// TIA Portal V21 export
// export: Created 2026-11-10T19:43:15.1099437Z, ExportSetting WithDefaults, DisplayName Totally Integrated Automation Portal, DisplayVersion V21 Update 3, DisplayName STEP 7 Professional, DisplayVersion V21 Update 3, DisplayName STEP 7 Safety, DisplayVersion V21, DisplayName Tech WebApplication, DisplayVersion V21, DisplayName WinCC Basic/Comfort/Advanced, DisplayVersion V21 Update 3, DisplayName WinCC Unified, DisplayVersion V21 Update 3
FUNCTION_BLOCK "FB_LadStruct"   // FB116, LAD
{ S7_Optimized_Access := 'TRUE' }
VERSION : 0.1
// stored: AutoNumber true, IsIECCheckEnabled false, IsRetainMemResEnabled false, MemoryReserve 100, SetENOAutomatically false, UDAEnableTagReadback false
   VAR_INPUT
      "a" : Bool;
      "b" : Bool;
      c : Bool;
      ia : Int;
   END_VAR
   VAR_OUTPUT
      q : Bool;
      q2 : Bool;
      io : Int;
      io2 : Int;
   END_VAR
   VAR
      ifc1 { S7_SetPoint := 'True'} : "FB_Iface";
      ton1 { S7_SetPoint := 'True'} : TON_TIME;
   END_VAR
BEGIN

REGION Network 1: Parallel branch
   // Branch with a second contact
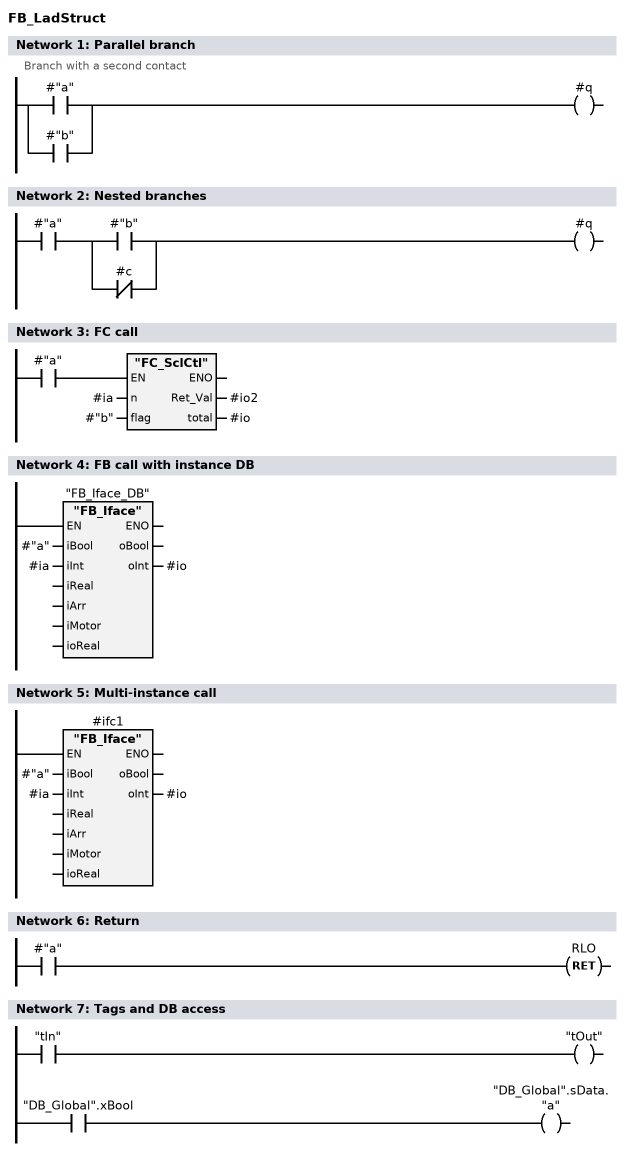
   RUNG wire#powerrail
      Contact( #"a" )
      wire#w1
      Coil( #q )
   END_RUNG
   RUNG wire#powerrail
      Contact( #"b" )
   END_RUNG wire#w1
   // the same network as SCL:
   #q := #"a" OR #"b";
END_REGION

REGION Network 2: Nested branches
   RUNG wire#powerrail
      Contact( #"a" )
      wire#w1
      Contact( #"b" )
      wire#w2
      Coil( #q )
   END_RUNG
   RUNG wire#w1
      I_Contact( #c )
   END_RUNG wire#w2
   // the same network as SCL:
   #q := #"a" AND (#"b" OR NOT #c);
END_REGION

REGION Network 3: FC call
   RUNG wire#powerrail
      Contact( #"a" )
      "FC_SclCtl"(n := #ia, flag := #"b", total => #io, Ret_Val => #io2)
   END_RUNG
   // the same network as SCL:
   IF #"a" THEN #io2 := "FC_SclCtl"(n := #ia, flag := #"b", total => #io); END_IF;
END_REGION

REGION Network 4: FB call with instance DB
   RUNG wire#powerrail
      "FB_Iface_DB"(iBool := #"a", iInt := #ia, oInt => #io, iReal :=, iArr :=, iMotor :=, oBool =>, ioReal :=)
   END_RUNG
   // the same network as SCL:
   "FB_Iface_DB"(iBool := #"a", iInt := #ia, oInt => #io);   // "FB_Iface"
END_REGION

REGION Network 5: Multi-instance call
   RUNG wire#powerrail
      #ifc1(iBool := #"a", iInt := #ia, oInt => #io, iReal :=, iArr :=, iMotor :=, oBool =>, ioReal :=)
   END_RUNG
   // the same network as SCL:
   #ifc1(iBool := #"a", iInt := #ia, oInt => #io);   // "FB_Iface"
END_REGION

REGION Network 6: Return
   IF #"a" THEN
       ENO := TRUE;
       RETURN;
   END_IF;
END_REGION

REGION Network 7: Tags and DB access
   RUNG wire#powerrail
      Contact( "tIn" )
      Coil( "tOut" )
   END_RUNG
   RUNG wire#powerrail
      Contact( "DB_Global".xBool )
      Coil( "DB_Global".sData."a" )
   END_RUNG
   // the same network as SCL:
   "tOut" := "tIn";
   "DB_Global".sData."a" := "DB_Global".xBool;
END_REGION
END_FUNCTION_BLOCK
